Universal Robots URScript: T015_zai-org_GLM-4.7-FP8_baseline_rep3.urscript

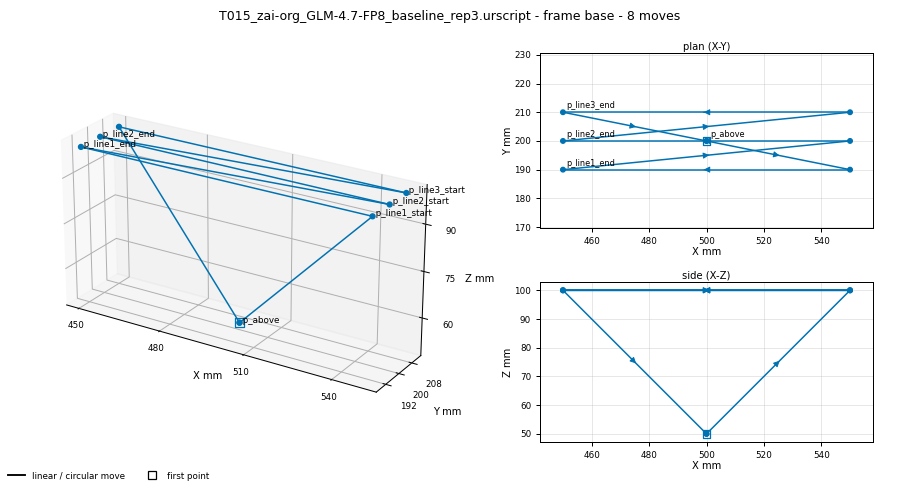
[picture p0: tool path of T015_zai-org_GLM-4.7-FP8_baseline_rep3.urscript in frame base, 8 of 10 moves have a stored position in this frame; points joined in program order, loops and branches not executed]
# URScript for Laser Marking Task T015
# Robot: UR5e, Mode: Fenced
# Payload: 0.6 kg

# Configuration
set_payload(0.6, [0.0, 0.0, 0.05])
set_tcp(p[0.0, 0.0, 0.0, 0.0, 0.0, 0.0])

# Global Variables
global home_joints = [0.0, -1.5708, 1.5708, -1.5708, -1.5708, 0.0]

# A6: Define Marking Fixture Frame
# Position: x=500mm, y=200mm, z=100mm, Rotation: Pointing down
global p_fixture = p[0.5, 0.2, 0.1, 0, 3.14159, 0]

# A3: Strict Laser Pointing - Define relative waypoints maintaining orientation
global p_above = pose_trans(p_fixture, p[0.0, 0.0, 0.05, 0.0, 0.0, 0.0])

# Line 1 (Y = -10mm)
global p_line1_start = pose_trans(p_fixture, p[-0.05, -0.01, 0.0, 0.0, 0.0, 0.0])
global p_line1_end   = pose_trans(p_fixture, p[ 0.05, -0.01, 0.0, 0.0, 0.0, 0.0])

# Line 2 (Y = 0mm)
global p_line2_start = pose_trans(p_fixture, p[-0.05,  0.0, 0.0, 0.0, 0.0, 0.0])
global p_line2_end   = pose_trans(p_fixture, p[ 0.05,  0.0, 0.0, 0.0, 0.0, 0.0])

# Line 3 (Y = 10mm)
global p_line3_start = pose_trans(p_fixture, p[-0.05,  0.01, 0.0, 0.0, 0.0, 0.0])
global p_line3_end   = pose_trans(p_fixture, p[ 0.05,  0.01, 0.0, 0.0, 0.0, 0.0])

# --- Motion Sequence ---

# 1. Move Joint: Home, 350.0 mm/s
movej(home_joints, a=1.4, v=0.35)

# 2. Move Linear: Above marking surface, 300.0 mm/s
movel(p_above, a=1.2, v=0.3)

# 3. Move Linear: Descend to marking height (Line 1 Start), 100.0 mm/s
movel(p_line1_start, a=0.5, v=0.1)

# 4. Move Linear: Mark line 1, 60.0 mm/s (A7: Laser Tool Activation)
set_digital_out(0, True)
movel(p_line1_end, a=0.2, v=0.06)
set_digital_out(0, False)

# 5. Move Linear: Step to line 2, 80.0 mm/s
movel(p_line2_start, a=0.5, v=0.08)

# 6. Move Linear: Mark line 2, 60.0 mm/s
set_digital_out(0, True)
movel(p_line2_end, a=0.2, v=0.06)
set_digital_out(0, False)

# 7. Move Linear: Step to line 3, 80.0 mm/s
movel(p_line3_start, a=0.5, v=0.08)

# 8. Move Linear: Mark line 3, 60.0 mm/s
set_digital_out(0, True)
movel(p_line3_end, a=0.2, v=0.06)
set_digital_out(0, False)

# 9. Move Linear: Retract to safety height, 200.0 mm/s
movel(p_above, a=0.5, v=0.2)

# 10. Move Joint: Return to Home, 350.0 mm/s
movej(home_joints, a=1.4, v=0.35)

# End of Program
